// TIA Portal V19 export
TYPE "EM06_Output"
   STRUCT
      Status : "EM_Output";
      DischargeActive : Bool;
      DrainActive : Bool;
      VacuumInterlock : Bool;
   END_STRUCT;
END_TYPE
